FUNCTION_BLOCK FB_KUKA_REF_1
VAR_INPUT
	KukaToPlc			:ST_KUKATOPLC;
	PlcToKuka			:ST_PLCTOKUKA;
END_VAR
VAR_OUTPUT

END_VAR
VAR_IN_OUT

END_VAR
VAR

END_VAR

;

END_FUNCTION_BLOCK

(* stored: Version 1.1.0.1, ProductVersion 3.1.4024.15
   POU FB_KUKA_REF_1: Id {0740f7e9-eb77-40d0-b8fe-21e80e7c9739}, SpecialFunc None *)
